(* IEC 61131-3 sources: Lasal-MCP/examples/SampleSource/5_ClassInputOutputSolution/Stations/MachineControl/MachineControl/Class/AlarmBuffer, 1 file *)

(* ---- AlarmBuffer.st ---- *)
(*!
<Class
	Name               = "AlarmBuffer"
	Revision           = "1.4"
	RealtimeTask       = "false"
	CyclicTask         = "true"
	DefCyclictime      = "10 ms"
	BackgroundTask     = "false"
	Sigmatek           = "false"
	OSInterface        = "false"
	HighPriority       = "false"
	Automatic          = "false"
	UpdateMode         = "Prescan"
	SharedCommandTable = "true"
	Objectsize         = "(536,120)"
	Comment            = "Class collects all Alarms and defines the switching conditions for the class OPMode.">
	<Channels>
	</Channels>
	<Dependencies>
		<Files>
			<File Path=".\Class\AlarmBuffer\AlarmBuffer_en.pdf"/>
			<File Path=".\Class\AlarmBuffer\AlarmBuffer_de.pdf"/>
		</Files>
	</Dependencies>
	<RevDoku>
		<Owner Company="Sigmatek"/>
		<Dokumentation Revision="1.4" Date="2016-10-10" Author="HubChr" Company="Sigmatek" Description="Added documentation pdfs."/>
		<Dokumentation Revision="1.3" Date="2016-09-27" Author="KaiAnd" Company="Sigmatek" Description="corrected class servers (deleted &quot;dead&quot; servers ond connected all from the base class)"/>
		<Dokumentation Revision="1.2" Date="2015-09-22" Company="Sigmatek" Description="Creation."/>
	</RevDoku>
	<Network Name="AlarmBuffer">
		<!-- List of Components in this network -->
		<Components>
			<Object
				Name       = "_base"
				Class      = "AlarmBufferBase"
				Position   = "(158,120)"
				Visualized = "true">
				<Channels>
					<Server Name="actOPMode"/>
					<Server Name="AlarmInfo"/>
					<Server Name="ClassSvr"/>
					<Server Name="GroupAutomatic"/>
					<Server Name="GroupError"/>
					<Server Name="GroupHoming"/>
					<Server Name="GroupInit"/>
					<Server Name="GroupManual"/>
					<Server Name="GroupSemiAuto"/>
					<Server Name="GroupSetup"/>
					<Server Name="GroupStop"/>
					<Server Name="QuitAll"/>
					<Server Name="QuitGroup"/>
					<Client Name="coOPModeConfig"/>
					<Client Name="No" Value="64"/>
					<Client Name="Parameter1"/>
					<Client Name="Parameter2"/>
				</Channels>
			</Object>
		</Components>
		<Comments>
		</Comments>
		<!-- List of Connections in this network -->
		<Connections>
			<Connection Source="this.ClassSvr" Destination="_base.ClassSvr" Vertices="(882,210),(710,210),"/>
			<Connection Source="this.QuitAll" Destination="_base.QuitAll" Vertices="(882,270),(710,270),"/>
			<Connection Source="_base.No" Destination="this.No" Vertices="(158,210),(38,210),"/>
			<Connection Source="_base.Parameter1" Destination="this.Parameter1" Vertices="(158,330),(38,330),"/>
			<Connection Source="_base.Parameter2" Destination="this.Parameter2" Vertices="(158,390),(38,390),"/>
			<Connection Source="_base.coOPModeConfig" Destination="this.coOPModeConfig" Vertices="(158,270),(38,270),"/>
			<Connection Source="this.QuitGroup" Destination="_base.QuitGroup" Vertices="(882,330),(710,330),"/>
			<Connection Source="this.actOPMode" Destination="_base.actOPMode" Vertices="(882,390),(710,390),"/>
			<Connection Source="this.GroupInit" Destination="_base.GroupInit" Vertices="(882,450),(710,450),"/>
			<Connection Source="this.GroupHoming" Destination="_base.GroupHoming" Vertices="(882,510),(710,510),"/>
			<Connection Source="this.GroupStop" Destination="_base.GroupStop" Vertices="(882,570),(710,570),"/>
			<Connection Source="this.GroupSetup" Destination="_base.GroupSetup" Vertices="(882,630),(710,630),"/>
			<Connection Source="this.GroupManual" Destination="_base.GroupManual" Vertices="(882,690),(710,690),"/>
			<Connection Source="this.GroupSemiAuto" Destination="_base.GroupSemiAuto" Vertices="(882,750),(710,750),"/>
			<Connection Source="this.GroupAutomatic" Destination="_base.GroupAutomatic" Vertices="(882,810),(710,810),"/>
			<Connection Source="this.GroupError" Destination="_base.GroupError" Vertices="(882,870),(710,870),"/>
		</Connections>
		<!-- Headerfiles -->
		<Options>
		</Options>
	</Network>
</Class>
*)
#pragma using AlarmBufferBase

AlarmBuffer : CLASS
: AlarmBufferBase
  //Servers:
  //Clients:
  //Variables:
  //Functions:

	FUNCTION VIRTUAL GLOBAL CyWork
		VAR_INPUT
			EAX 	: UDINT;
		END_VAR
		VAR_OUTPUT
			state (EAX) 	: UDINT;
		END_VAR;

	FUNCTION VIRTUAL OPModeChange
		VAR_INPUT
			eActOPMode 	: t_e_OPMode;
			eNewOPMode 	: t_e_OPMode;
		END_VAR
		VAR_OUTPUT
			bOK 	: BOOL;
		END_VAR;

	FUNCTION VIRTUAL OPModeActive
		VAR_INPUT
			eActOPMode 	: t_e_OPMode;
		END_VAR
		VAR_OUTPUT
			eNewOPMode 	: t_e_OPMode;
		END_VAR;
  //Tables:
	FUNCTION @STD
		VAR_OUTPUT
			ret_code	: CONFSTATES;
		END_VAR;
	FUNCTION GLOBAL TAB @CT_;
END_CLASS;

FUNCTION VIRTUAL AlarmBuffer::OPModeChange
	VAR_INPUT
		eActOPMode 	: t_e_OPMode;
		eNewOPMode 	: t_e_OPMode;
	END_VAR
	VAR_OUTPUT
		bOK 	: BOOL;
	END_VAR

  bOK := true;

  //*****************************************************************************
  //** UNTERSCHEIDUNG FÜR NEUEN BETRIEBSMODUS                                  **
  //*****************************************************************************

  // je nachdem in welchen Betriebsmodus gewechselt werden soll, müssen die
  // Alarme geprüft werden. Ein Alarm kann einen Wechsel in einen anderen
  // Betriebsmodus verhindern.
  // aktueller Betriebsmodus = Manual
  // neuer Betriebsmodus = Automatik
  // Alarm mit der Gruppe SemiAutomatik aktiv
  // => Umschalten wird verhindert

  case eNewOPMode of

    // Betriebsart Init
    //***************************************************************************
    OPMode_Init:

      // in diesen Betriebsmodus kann immer gewechselt werden,
      // egal welche Alarme aktiv sind.

    // Betriebsart Homing
    //***************************************************************************
    OPMode_Homing:

      // in diesen Betriebsmodus kann immer gewechselt werden,
      // egal welche Alarme aktiv sind.

    // Betriebsmodus Stop
    //***************************************************************************
    OPMode_Stop:

      // in diesen Betriebsmodus kann immer gewechselt werden,
      // egal welche Alarme aktiv sind.

    // Betriebsmodus Manual + Setup
    //***************************************************************************
    OPMode_Manual, OPMode_Setup:

      // Prüfen ob Alarm der Gruppe Stop aktiv ist
      //------------------------------------------------------
      if sOPModeAlarm.udOPModeStop then
        bOK := false;
      end_if;

    // Betriebsmodus SemiAutomatic
    //***************************************************************************
    OPMode_SemiAuto:

      // Prüfen ob Alarm der Gruppe Stop oder Manual aktiv ist
      //------------------------------------------------------
      if  sOPModeAlarm.udOPModeStop |
          sOPModeAlarm.udOPModeManual then
        bOK := false;
      end_if;

    // Betriebsmodus Automatic
    //***************************************************************************
    OPMode_Automatic:

      // Prüfen ob Alarm der Gruppe Stop, Manual oder Halbautomatik aktiv ist
      //------------------------------------------------------
      if  sOPModeAlarm.udOPModeStop |
          sOPModeAlarm.udOPModeManual |
          sOPModeAlarm.udOPModeSemiAuto then
        bOK := false;
      end_if;

    // Betriebsmodus Error
    //***************************************************************************
    OPMode_Error:

      // in diesen Betriebsmodus kann immer gewechselt werden,
      // egal welche Alarme aktiv sind.

    // nicht unterstützer Betriebsmodus
    //***************************************************************************
    else
      TRACE("AlarmBuffer::OPModeChange(): nicht unterstützter Betriebsmodus aktiv");
      bOK := false;

  end_case;

END_FUNCTION

FUNCTION VIRTUAL AlarmBuffer::OPModeActive
	VAR_INPUT
		eActOPMode 	: t_e_OPMode;
	END_VAR
	VAR_OUTPUT
		eNewOPMode 	: t_e_OPMode;
	END_VAR

  // Rückgabewert initialisieren
  // => kein Wechsel Betriebsmodus
  eNewOPMode := eActOPMode;

  //*****************************************************************************
  //** FÜR DEN AKTUELLEN BETRIEBSMODUS ALARME PRÜFEN                           **
  //*****************************************************************************

  // Die OPMode-Gruppe eines Alarmes definiert, in welchen Betriebsmodus
  // gewechselt werden muss, wenn der Alarm auftritt. Dabei wird der Modus
  // Automatik am höchsten bewertet, der Modus Manual am niedrigsten.
  // Tritt daher im Modus SemiAuto ein Alarm der Gruppe Automatik auf, so
  // wird nicht gewechselt.

  case eActOPMode of

    // Betriebsmodus Init
    //***************************************************************************
    OPMode_Init:

      // im Betriebsmodus Init können Alarme auftreten, ohne dass der Modus
      // gewechselt werden muss.

    // Betriebsmodus Stop
    //***************************************************************************
    OPMode_Stop:

      // im Betriebsmodus Stop können Alarme auftreten, ohne dass der Modus
      // gewechselt werden muss.

    // Betriebsmodus Manual + Setup
    //***************************************************************************
    OPMode_Manual, OPMode_Setup:

      // Prüfen ob Alarm der Gruppe Stop aktiv ist
      //---------------------------------------------
      if sOPModeAlarm.udOPModeStop then
        eNewOPMode := OPMode_Stop;
      end_if;

      // Prüfen ob Alarm der Gruppe Error aktiv ist
      // --------------------------------------------
      if sOPModeAlarm.udOPModeError then
        eNewOPMode := OPMode_Error;
      end_if;

    // Betriebsmodus SemiAuto
    //***************************************************************************
    OPMode_SemiAuto:

      // Prüfen ob Alarm der Gruppe Stop aktiv ist
      //---------------------------------------------
      if sOPModeAlarm.udOPModeStop then
        eNewOPMode := OPMode_Stop;

      // Prüfen ob Alarm der Gruppe Manual aktiv ist
      //---------------------------------------------
      elsif sOPModeAlarm.udOPModeManual then
        eNewOPMode := OPMode_Manual;

      end_if;

    // Betriebsmodus Automatic
    //***************************************************************************
    OPMode_Automatic:

      // Prüfen ob Alarm der Gruppe Stop aktiv ist
      //---------------------------------------------
      if sOPModeAlarm.udOPModeStop then
        eNewOPMode := OPMode_Stop;

      // Prüfen ob Alarm der Gruppe Manual aktiv ist
      //---------------------------------------------
      elsif sOPModeAlarm.udOPModeManual then
        eNewOPMode := OPMode_Manual;

      // Prüfen ob Alarm der Gruppe SemiAuto aktiv ist
      //----------------------------------------------
      elsif sOPModeAlarm.udOPModeSemiAuto then
        eNewOPMode := OPMode_SemiAuto;

      end_if;

    // nicht unterstützer Betriebsmodus
    //***************************************************************************
    else
      TRACE("AlarmBuffer::CheckAlarm(): nicht unterstützter Betriebsmodus aktiv");
      eActOPMode := OPMode_Stop;

  end_case;

END_FUNCTION

FUNCTION VIRTUAL GLOBAL AlarmBuffer::CyWork
	VAR_INPUT
		EAX 	: UDINT;
	END_VAR
	VAR_OUTPUT
		state (EAX) 	: UDINT;
	END_VAR

  // aktive Alarme auf den Server darstellen
  GroupInit       := sOPModeAlarm.udOPModeInit;
  GroupHoming     := sOPModeAlarm.udOPModeHoming;
  GroupStop       := sOPModeAlarm.udOPModeStop;
  GroupSetup      := sOPModeAlarm.udOPModeSetup;
  GroupManual     := sOPModeAlarm.udOPModeManual;
  GroupSemiAuto   := sOPModeAlarm.udOPModeSemiAuto;
  GroupAutomatic  := sOPModeAlarm.udOPModeAutomatic;
  GroupError      := sOPModeAlarm.udOPModeError;

	state := READY;

END_FUNCTION
